(* IEC 61131-3 sources: plc-st-coding-agent/progress/evidence/f14_v13_self_20261113/jobs/custom_deepseek-v4pro (part 4) *)

(* ---- public-medium-02.raw_candidate_01.st ---- *)
TYPE ST_AnalogChannel :
STRUCT
    enable : BOOL;
    hiLIM : REAL;
    loLIM : REAL;
    bipolar : BOOL;
    measuringMode : INT;
    retVal : WORD;
    outputValue : REAL;
END_STRUCT
END_TYPE

(* ENGINEERING_CONTRACT
   Loop count: count limited to 0..min(array lengths); ordinal start at each array lower bound (PUB001).
   channels[].retVal: activated on enabled scan; invalid mode -> 16#8001, invalid limits -> 16#8002,
   success -> 0 (PUB006, PUB007, PUB008).
   channels[].outputValue: written only on successful conversion; mode 0 linear scaling,
   mode 1 /10, mode 2 /100 (PUB003, PUB004, PUB005).
   Disabled channels retain prior retVal/outputValue (unspecified retention interpretation).
*)

(* CONTRACT_RULES [] *)

FUNCTION_BLOCK AnalogBatchProcessing
VAR_INPUT
    count : DINT;
END_VAR
VAR_IN_OUT
    analogValues : ARRAY[*] OF INT;
    channels : ARRAY[*] OF ST_AnalogChannel;
END_VAR
VAR
    local_i : DINT;
    local_n : DINT;
    local_analog_idx : DINT;
    local_channel_idx : DINT;
    local_raw : INT;
    local_mode : INT;
    local_min_len : DINT;
    local_ch_len : DINT;
    local_raw_min : REAL;
    local_raw_max : REAL;
    local_span_raw : REAL;
    local_ratio : REAL;
END_VAR

local_n := count;
IF local_n < 0 THEN
    local_n := 0;
END_IF;

local_min_len := UPPER_BOUND(analogValues, 1) - LOWER_BOUND(analogValues, 1) + 1;
local_ch_len := UPPER_BOUND(channels, 1) - LOWER_BOUND(channels, 1) + 1;
IF local_min_len > local_ch_len THEN
    local_min_len := local_ch_len;
END_IF;
IF local_n > local_min_len THEN
    local_n := local_min_len;
END_IF;

IF local_n > 0 THEN
    FOR local_i := 0 TO local_n - 1 DO
        local_analog_idx := LOWER_BOUND(analogValues, 1) + local_i;
        local_channel_idx := LOWER_BOUND(channels, 1) + local_i;

        IF channels[local_channel_idx].enable THEN
            local_mode := channels[local_channel_idx].measuringMode;

            IF (local_mode <> 0) AND (local_mode <> 1) AND (local_mode <> 2) THEN
                channels[local_channel_idx].retVal := 16#8001;
                (* skip conversion: outputValue unchanged *)
            ELSIF channels[local_channel_idx].hiLIM <= channels[local_channel_idx].loLIM THEN
                channels[local_channel_idx].retVal := 16#8002;
                (* skip conversion: outputValue unchanged *)
            ELSE
                channels[local_channel_idx].retVal := 0;
                CASE local_mode OF
                    0:
                        local_raw := analogValues[local_analog_idx];
                        IF channels[local_channel_idx].bipolar THEN
                            local_raw_min := -27648.0;
                            local_raw_max := 27648.0;
                        ELSE
                            local_raw_min := 0.0;
                            local_raw_max := 27648.0;
                        END_IF;

                        local_span_raw := local_raw_max - local_raw_min;
                        local_ratio := (TO_REAL(local_raw) - local_raw_min) / local_span_raw;
                        channels[local_channel_idx].outputValue := channels[local_channel_idx].loLIM
                            + local_ratio * (channels[local_channel_idx].hiLIM - channels[local_channel_idx].loLIM);

                    1:
                        channels[local_channel_idx].outputValue := TO_REAL(analogValues[local_analog_idx]) / 10.0;

                    2:
                        channels[local_channel_idx].outputValue := TO_REAL(analogValues[local_analog_idx]) / 100.0;
                END_CASE;
            END_IF;
        ELSE
            (* disabled: no writes to retVal or outputValue *)
        END_IF;
    END_FOR;
END_IF;

(* ---- public-medium-02.raw_candidate_02.st ---- *)
TYPE ST_AnalogChannel :
STRUCT
    enable : BOOL;
    hiLIM : REAL;
    loLIM : REAL;
    bipolar : BOOL;
    measuringMode : INT;
    retVal : WORD;
    outputValue : REAL;
END_STRUCT
END_TYPE;

(* ENGINEERING_CONTRACT
   Loop count: count limited to 0..min(array lengths); ordinal start at each array lower bound (PUB001).
   channels[].retVal: activated on enabled scan; invalid mode -> 16#8001, invalid limits -> 16#8002,
   success -> 0 (PUB006, PUB007, PUB008).
   channels[].outputValue: written only on successful conversion; mode 0 linear scaling,
   mode 1 /10, mode 2 /100 (PUB003, PUB004, PUB005).
   Disabled channels retain prior retVal/outputValue (unspecified retention interpretation).
*)

(* CONTRACT_RULES [] *)

FUNCTION_BLOCK AnalogBatchProcessing
VAR_INPUT
    count : DINT;
END_VAR
VAR_IN_OUT
    analogValues : ARRAY[*] OF INT;
    channels : ARRAY[*] OF ST_AnalogChannel;
END_VAR
VAR
    local_i : DINT;
    local_n : DINT;
    local_analog_idx : DINT;
    local_channel_idx : DINT;
    local_raw : INT;
    local_mode : INT;
    local_min_len : DINT;
    local_ch_len : DINT;
    local_raw_min : REAL;
    local_raw_max : REAL;
    local_span_raw : REAL;
    local_ratio : REAL;
END_VAR

local_n := count;
IF local_n < 0 THEN
    local_n := 0;
END_IF;

local_min_len := UPPER_BOUND(analogValues, 1) - LOWER_BOUND(analogValues, 1) + 1;
local_ch_len := UPPER_BOUND(channels, 1) - LOWER_BOUND(channels, 1) + 1;
IF local_min_len > local_ch_len THEN
    local_min_len := local_ch_len;
END_IF;
IF local_n > local_min_len THEN
    local_n := local_min_len;
END_IF;

IF local_n > 0 THEN
    FOR local_i := 0 TO local_n - 1 DO
        local_analog_idx := LOWER_BOUND(analogValues, 1) + local_i;
        local_channel_idx := LOWER_BOUND(channels, 1) + local_i;

        IF channels[local_channel_idx].enable THEN
            local_mode := channels[local_channel_idx].measuringMode;

            IF (local_mode <> 0) AND (local_mode <> 1) AND (local_mode <> 2) THEN
                channels[local_channel_idx].retVal := 16#8001;
                (* skip conversion: outputValue unchanged *)
            ELSIF channels[local_channel_idx].hiLIM <= channels[local_channel_idx].loLIM THEN
                channels[local_channel_idx].retVal := 16#8002;
                (* skip conversion: outputValue unchanged *)
            ELSE
                channels[local_channel_idx].retVal := 0;
                CASE local_mode OF
                    0:
                        local_raw := analogValues[local_analog_idx];
                        IF channels[local_channel_idx].bipolar THEN
                            local_raw_min := -27648.0;
                            local_raw_max := 27648.0;
                        ELSE
                            local_raw_min := 0.0;
                            local_raw_max := 27648.0;
                        END_IF;

                        local_span_raw := local_raw_max - local_raw_min;
                        local_ratio := (TO_REAL(local_raw) - local_raw_min) / local_span_raw;
                        channels[local_channel_idx].outputValue := channels[local_channel_idx].loLIM
                            + local_ratio * (channels[local_channel_idx].hiLIM - channels[local_channel_idx].loLIM);

                    1:
                        channels[local_channel_idx].outputValue := TO_REAL(analogValues[local_analog_idx]) / 10.0;

                    2:
                        channels[local_channel_idx].outputValue := TO_REAL(analogValues[local_analog_idx]) / 100.0;
                END_CASE;
            END_IF;
        ELSE
            (* disabled: no writes to retVal or outputValue *)
        END_IF;
    END_FOR;
END_IF;

END_FUNCTION_BLOCK

(* ---- public-medium-02.raw_candidate_03.st ---- *)
TYPE ST_AnalogChannel :
STRUCT
    enable : BOOL;
    hiLIM : REAL;
    loLIM : REAL;
    bipolar : BOOL;
    measuringMode : INT;
    retVal : WORD;
    outputValue : REAL;
END_STRUCT
END_TYPE

(* ENGINEERING_CONTRACT
   Loop count: count limited to 0..min(array lengths); ordinal start at each array lower bound (PUB001).
   channels[].retVal: activated on enabled scan; invalid mode -> 16#8001, invalid limits -> 16#8002,
   success -> 0 (PUB006, PUB007, PUB008).
   channels[].outputValue: written only on successful conversion; mode 0 linear scaling,
   mode 1 /10, mode 2 /100 (PUB003, PUB004, PUB005).
   Disabled channels retain prior retVal/outputValue (unspecified retention interpretation).
*)

(* CONTRACT_RULES [] *)

FUNCTION_BLOCK AnalogBatchProcessing
VAR_INPUT
    count : DINT;
END_VAR
VAR_IN_OUT
    analogValues : ARRAY[*] OF INT;
    channels : ARRAY[*] OF ST_AnalogChannel;
END_VAR
VAR
    local_i : DINT;
    local_n : DINT;
    local_analog_idx : DINT;
    local_channel_idx : DINT;
    local_raw : INT;
    local_mode : INT;
    local_min_len : DINT;
    local_ch_len : DINT;
    local_raw_min : REAL;
    local_raw_max : REAL;
    local_span_raw : REAL;
    local_ratio : REAL;
END_VAR

local_n := count;
IF local_n < 0 THEN
    local_n := 0;
END_IF;

local_min_len := UPPER_BOUND(analogValues, 1) - LOWER_BOUND(analogValues, 1) + 1;
local_ch_len := UPPER_BOUND(channels, 1) - LOWER_BOUND(channels, 1) + 1;
IF local_min_len > local_ch_len THEN
    local_min_len := local_ch_len;
END_IF;
IF local_n > local_min_len THEN
    local_n := local_min_len;
END_IF;

IF local_n > 0 THEN
    FOR local_i := 0 TO local_n - 1 DO
        local_analog_idx := LOWER_BOUND(analogValues, 1) + local_i;
        local_channel_idx := LOWER_BOUND(channels, 1) + local_i;

        IF channels[local_channel_idx].enable THEN
            local_mode := channels[local_channel_idx].measuringMode;

            IF (local_mode <> 0) AND (local_mode <> 1) AND (local_mode <> 2) THEN
                channels[local_channel_idx].retVal := 16#8001;
                (* skip conversion: outputValue unchanged *)
            ELSIF channels[local_channel_idx].hiLIM <= channels[local_channel_idx].loLIM THEN
                channels[local_channel_idx].retVal := 16#8002;
                (* skip conversion: outputValue unchanged *)
            ELSE
                channels[local_channel_idx].retVal := 0;
                CASE local_mode OF
                    0:
                        local_raw := analogValues[local_analog_idx];
                        IF channels[local_channel_idx].bipolar THEN
                            local_raw_min := -27648.0;
                            local_raw_max := 27648.0;
                        ELSE
                            local_raw_min := 0.0;
                            local_raw_max := 27648.0;
                        END_IF;

                        local_span_raw := local_raw_max - local_raw_min;
                        local_ratio := (TO_REAL(local_raw) - local_raw_min) / local_span_raw;
                        channels[local_channel_idx].outputValue := channels[local_channel_idx].loLIM
                            + local_ratio * (channels[local_channel_idx].hiLIM - channels[local_channel_idx].loLIM);

                    1:
                        channels[local_channel_idx].outputValue := TO_REAL(analogValues[local_analog_idx]) / 10.0;

                    2:
                        channels[local_channel_idx].outputValue := TO_REAL(analogValues[local_analog_idx]) / 100.0;
                END_CASE;
            END_IF;
        ELSE
            (* disabled: no writes to retVal or outputValue *)
        END_IF;
    END_FOR;
END_IF;

END_FUNCTION_BLOCK

(* ---- public-medium-03.candidate_01.st ---- *)
(* ENGINEERING_CONTRACT
- average: stored LREAL; updated on valid acquisition; reset or invalid window clears it to 0.0.
- windowSizeReached: FALSE until count >= windowSize; retained until reset or invalid window.
- error/status: combinational invalid windowSize (1..100 inclusive); otherwise clear/zero.
- Priority: invalid window first, reset second, acquisition last (reset priority chosen).
- cyclicExecution TRUE ignores trigger edges for extra samples (PUB001/2).
- trigger edge is evaluated only from previous scan raw trigger state.
- Same-scan: validate window, detect window-size change, reset, acquire, update average.
*)
(* CONTRACT_RULES [] *)
FUNCTION_BLOCK FB
VAR_INPUT
    cyclicExecution : BOOL;
    trigger : BOOL;
    value : LREAL;
    windowSize : INT;
    reset : BOOL;
END_VAR
VAR_OUTPUT
    average : LREAL;
    windowSizeReached : BOOL;
    error : BOOL;
    status : WORD;
END_VAR
VAR
    tmp_buffer : ARRAY[0..99] OF LREAL;
    tmp_count : INT := 0;
    tmp_index : INT := 0;
    tmp_sum : LREAL := 0.0;
    tmp_previousTrigger : BOOL := FALSE;
    tmp_windowSize : INT := 0;
END_VAR

IF (windowSize < 1) OR (windowSize > 100) THEN
    error := TRUE;
    status := WORD#16#8200;
    windowSizeReached := FALSE;
    average := 0.0;
    tmp_count := 0;
    tmp_index := 0;
    tmp_sum := 0.0;
    tmp_windowSize := windowSize;
ELSE
    error := FALSE;
    status := WORD#16#0000;

    IF tmp_windowSize <> windowSize THEN
        tmp_count := 0;
        tmp_index := 0;
        tmp_sum := 0.0;
        windowSizeReached := FALSE;
        average := 0.0;
        tmp_windowSize := windowSize;
    END_IF;

    IF reset THEN
        tmp_count := 0;
        tmp_index := 0;
        tmp_sum := 0.0;
        windowSizeReached := FALSE;
        average := 0.0;
    ELSE
        IF cyclicExecution OR (trigger AND NOT tmp_previousTrigger) THEN
            IF tmp_count < windowSize THEN
                tmp_count := tmp_count + 1;
                tmp_sum := tmp_sum + value;
                tmp_buffer[tmp_index] := value;
                tmp_index := tmp_index + 1;
                IF tmp_index >= windowSize THEN
                    tmp_index := 0;
                END_IF;
            ELSE
                tmp_sum := tmp_sum - tmp_buffer[tmp_index] + value;
                tmp_buffer[tmp_index] := value;
                tmp_index := tmp_index + 1;
                IF tmp_index >= windowSize THEN
                    tmp_index := 0;
                END_IF;
            END_IF;

            average := tmp_sum / INT_TO_LREAL(tmp_count);
            windowSizeReached := tmp_count >= windowSize;
        END_IF;
    END_IF;
END_IF;

tmp_previousTrigger := trigger;

(* ---- public-medium-03.candidate_02.st ---- *)
(* ENGINEERING_CONTRACT
- average: stored LREAL; updated on valid acquisition; reset or invalid window clears it to 0.0.
- windowSizeReached: FALSE until count >= windowSize; retained until reset or invalid window.
- error/status: combinational invalid windowSize (1..100 inclusive); otherwise clear/zero.
- Priority: invalid window first, reset second, acquisition last (reset priority chosen).
- cyclicExecution TRUE ignores trigger edges for extra samples (PUB001/2).
- trigger edge is evaluated only from previous scan raw trigger state.
- Same-scan: validate window, detect window-size change, reset, acquire, update average.
*)
(* CONTRACT_RULES [] *)
FUNCTION_BLOCK FB
VAR_INPUT
    cyclicExecution : BOOL;
    trigger : BOOL;
    value : LREAL;
    windowSize : INT;
    reset : BOOL;
END_VAR
VAR_OUTPUT
    average : LREAL;
    windowSizeReached : BOOL;
    error : BOOL;
    status : WORD;
END_VAR
VAR
    tmp_buffer : ARRAY[0..99] OF LREAL;
    tmp_count : INT := 0;
    tmp_index : INT := 0;
    tmp_sum : LREAL := 0.0;
    tmp_previousTrigger : BOOL := FALSE;
    tmp_windowSize : INT := 0;
END_VAR

IF (windowSize < 1) OR (windowSize > 100) THEN
    error := TRUE;
    status := WORD#16#8200;
    windowSizeReached := FALSE;
    average := 0.0;
    tmp_count := 0;
    tmp_index := 0;
    tmp_sum := 0.0;
    tmp_windowSize := windowSize;
ELSE
    error := FALSE;
    status := WORD#16#0000;

    IF tmp_windowSize <> windowSize THEN
        tmp_count := 0;
        tmp_index := 0;
        tmp_sum := 0.0;
        windowSizeReached := FALSE;
        average := 0.0;
        tmp_windowSize := windowSize;
    END_IF;

    IF reset THEN
        tmp_count := 0;
        tmp_index := 0;
        tmp_sum := 0.0;
        windowSizeReached := FALSE;
        average := 0.0;
    ELSE
        IF cyclicExecution OR (trigger AND NOT tmp_previousTrigger) THEN
            IF tmp_count < windowSize THEN
                tmp_count := tmp_count + 1;
                tmp_sum := tmp_sum + value;
                tmp_buffer[tmp_index] := value;
                tmp_index := tmp_index + 1;
                IF tmp_index >= windowSize THEN
                    tmp_index := 0;
                END_IF;
            ELSE
                tmp_sum := tmp_sum - tmp_buffer[tmp_index] + value;
                tmp_buffer[tmp_index] := value;
                tmp_index := tmp_index + 1;
                IF tmp_index >= windowSize THEN
                    tmp_index := 0;
                END_IF;
            END_IF;

            average := tmp_sum / INT_TO_LREAL(tmp_count);
            windowSizeReached := tmp_count >= windowSize;
        END_IF;
    END_IF;
END_IF;

tmp_previousTrigger := trigger;
END_FUNCTION_BLOCK

(* ---- public-medium-03.patch_base_02.st ---- *)
(* ENGINEERING_CONTRACT
- average: stored LREAL; updated on valid acquisition; reset or invalid window clears it to 0.0.
- windowSizeReached: FALSE until count >= windowSize; retained until reset or invalid window.
- error/status: combinational invalid windowSize (1..100 inclusive); otherwise clear/zero.
- Priority: invalid window first, reset second, acquisition last (reset priority chosen).
- cyclicExecution TRUE ignores trigger edges for extra samples (PUB001/2).
- trigger edge is evaluated only from previous scan raw trigger state.
- Same-scan: validate window, detect window-size change, reset, acquire, update average.
*)
(* CONTRACT_RULES [] *)
FUNCTION_BLOCK FB
VAR_INPUT
    cyclicExecution : BOOL;
    trigger : BOOL;
    value : LREAL;
    windowSize : INT;
    reset : BOOL;
END_VAR
VAR_OUTPUT
    average : LREAL;
    windowSizeReached : BOOL;
    error : BOOL;
    status : WORD;
END_VAR
VAR
    tmp_buffer : ARRAY[0..99] OF LREAL;
    tmp_count : INT := 0;
    tmp_index : INT := 0;
    tmp_sum : LREAL := 0.0;
    tmp_previousTrigger : BOOL := FALSE;
    tmp_windowSize : INT := 0;
END_VAR

IF (windowSize < 1) OR (windowSize > 100) THEN
    error := TRUE;
    status := WORD#16#8200;
    windowSizeReached := FALSE;
    average := 0.0;
    tmp_count := 0;
    tmp_index := 0;
    tmp_sum := 0.0;
    tmp_windowSize := windowSize;
ELSE
    error := FALSE;
    status := WORD#16#0000;

    IF tmp_windowSize <> windowSize THEN
        tmp_count := 0;
        tmp_index := 0;
        tmp_sum := 0.0;
        windowSizeReached := FALSE;
        average := 0.0;
        tmp_windowSize := windowSize;
    END_IF;

    IF reset THEN
        tmp_count := 0;
        tmp_index := 0;
        tmp_sum := 0.0;
        windowSizeReached := FALSE;
        average := 0.0;
    ELSE
        IF cyclicExecution OR (trigger AND NOT tmp_previousTrigger) THEN
            IF tmp_count < windowSize THEN
                tmp_count := tmp_count + 1;
                tmp_sum := tmp_sum + value;
                tmp_buffer[tmp_index] := value;
                tmp_index := tmp_index + 1;
                IF tmp_index >= windowSize THEN
                    tmp_index := 0;
                END_IF;
            ELSE
                tmp_sum := tmp_sum - tmp_buffer[tmp_index] + value;
                tmp_buffer[tmp_index] := value;
                tmp_index := tmp_index + 1;
                IF tmp_index >= windowSize THEN
                    tmp_index := 0;
                END_IF;
            END_IF;

            average := tmp_sum / INT_TO_LREAL(tmp_count);
            windowSizeReached := tmp_count >= windowSize;
        END_IF;
    END_IF;
END_IF;

tmp_previousTrigger := trigger;

(* ---- public-medium-03.raw_candidate_01.st ---- *)
(* ENGINEERING_CONTRACT
- average: stored LREAL; updated on valid acquisition; reset or invalid window clears it to 0.0.
- windowSizeReached: FALSE until count >= windowSize; retained until reset or invalid window.
- error/status: combinational invalid windowSize (1..100 inclusive); otherwise clear/zero.
- Priority: invalid window first, reset second, acquisition last (reset priority chosen).
- cyclicExecution TRUE ignores trigger edges for extra samples (PUB001/2).
- trigger edge is evaluated only from previous scan raw trigger state.
- Same-scan: validate window, detect window-size change, reset, acquire, update average.
*)
(* CONTRACT_RULES [] *)
FUNCTION_BLOCK FB
VAR_INPUT
    cyclicExecution : BOOL;
    trigger : BOOL;
    value : LREAL;
    windowSize : INT;
    reset : BOOL;
END_VAR
VAR_OUTPUT
    average : LREAL;
    windowSizeReached : BOOL;
    error : BOOL;
    status : WORD;
END_VAR
VAR
    tmp_buffer : ARRAY[0..99] OF LREAL;
    tmp_count : INT := 0;
    tmp_index : INT := 0;
    tmp_sum : LREAL := 0.0;
    tmp_previousTrigger : BOOL := FALSE;
    tmp_windowSize : INT := 0;
END_VAR

IF (windowSize < 1) OR (windowSize > 100) THEN
    error := TRUE;
    status := WORD#16#8200;
    windowSizeReached := FALSE;
    average := 0.0;
    tmp_count := 0;
    tmp_index := 0;
    tmp_sum := 0.0;
    tmp_windowSize := windowSize;
ELSE
    error := FALSE;
    status := WORD#16#0000;

    IF tmp_windowSize <> windowSize THEN
        tmp_count := 0;
        tmp_index := 0;
        tmp_sum := 0.0;
        windowSizeReached := FALSE;
        average := 0.0;
        tmp_windowSize := windowSize;
    END_IF;

    IF reset THEN
        tmp_count := 0;
        tmp_index := 0;
        tmp_sum := 0.0;
        windowSizeReached := FALSE;
        average := 0.0;
    ELSE
        IF cyclicExecution OR (trigger AND NOT tmp_previousTrigger) THEN
            IF tmp_count < windowSize THEN
                tmp_count := tmp_count + 1;
                tmp_sum := tmp_sum + value;
                tmp_buffer[tmp_index] := value;
                tmp_index := tmp_index + 1;
                IF tmp_index >= windowSize THEN
                    tmp_index := 0;
                END_IF;
            ELSE
                tmp_sum := tmp_sum - tmp_buffer[tmp_index] + value;
                tmp_buffer[tmp_index] := value;
                tmp_index := tmp_index + 1;
                IF tmp_index >= windowSize THEN
                    tmp_index := 0;
                END_IF;
            END_IF;

            average := tmp_sum / INT_TO_LREAL(tmp_count);
            windowSizeReached := tmp_count >= windowSize;
        END_IF;
    END_IF;
END_IF;

tmp_previousTrigger := trigger;

(* ---- public-medium-03.raw_candidate_02.st ---- *)
(* ENGINEERING_CONTRACT
- average: stored LREAL; updated on valid acquisition; reset or invalid window clears it to 0.0.
- windowSizeReached: FALSE until count >= windowSize; retained until reset or invalid window.
- error/status: combinational invalid windowSize (1..100 inclusive); otherwise clear/zero.
- Priority: invalid window first, reset second, acquisition last (reset priority chosen).
- cyclicExecution TRUE ignores trigger edges for extra samples (PUB001/2).
- trigger edge is evaluated only from previous scan raw trigger state.
- Same-scan: validate window, detect window-size change, reset, acquire, update average.
*)
(* CONTRACT_RULES [] *)
FUNCTION_BLOCK FB
VAR_INPUT
    cyclicExecution : BOOL;
    trigger : BOOL;
    value : LREAL;
    windowSize : INT;
    reset : BOOL;
END_VAR
VAR_OUTPUT
    average : LREAL;
    windowSizeReached : BOOL;
    error : BOOL;
    status : WORD;
END_VAR
VAR
    tmp_buffer : ARRAY[0..99] OF LREAL;
    tmp_count : INT := 0;
    tmp_index : INT := 0;
    tmp_sum : LREAL := 0.0;
    tmp_previousTrigger : BOOL := FALSE;
    tmp_windowSize : INT := 0;
END_VAR

IF (windowSize < 1) OR (windowSize > 100) THEN
    error := TRUE;
    status := WORD#16#8200;
    windowSizeReached := FALSE;
    average := 0.0;
    tmp_count := 0;
    tmp_index := 0;
    tmp_sum := 0.0;
    tmp_windowSize := windowSize;
ELSE
    error := FALSE;
    status := WORD#16#0000;

    IF tmp_windowSize <> windowSize THEN
        tmp_count := 0;
        tmp_index := 0;
        tmp_sum := 0.0;
        windowSizeReached := FALSE;
        average := 0.0;
        tmp_windowSize := windowSize;
    END_IF;

    IF reset THEN
        tmp_count := 0;
        tmp_index := 0;
        tmp_sum := 0.0;
        windowSizeReached := FALSE;
        average := 0.0;
    ELSE
        IF cyclicExecution OR (trigger AND NOT tmp_previousTrigger) THEN
            IF tmp_count < windowSize THEN
                tmp_count := tmp_count + 1;
                tmp_sum := tmp_sum + value;
                tmp_buffer[tmp_index] := value;
                tmp_index := tmp_index + 1;
                IF tmp_index >= windowSize THEN
                    tmp_index := 0;
                END_IF;
            ELSE
                tmp_sum := tmp_sum - tmp_buffer[tmp_index] + value;
                tmp_buffer[tmp_index] := value;
                tmp_index := tmp_index + 1;
                IF tmp_index >= windowSize THEN
                    tmp_index := 0;
                END_IF;
            END_IF;

            average := tmp_sum / INT_TO_LREAL(tmp_count);
            windowSizeReached := tmp_count >= windowSize;
        END_IF;
    END_IF;
END_IF;

tmp_previousTrigger := trigger;
END_FUNCTION_BLOCK

(* ---- public-medium-04.candidate_01.st ---- *)
FUNCTION_BLOCK FB_TemperatureControl
VAR_INPUT
    TemperatureSensorInput : REAL;
    SetTemperature : REAL;
END_VAR
VAR_OUTPUT
    CurrentTemperature : REAL;
    SetTempDisplay : REAL;
    HeaterStatus : BOOL;
    OverheatProtection : BOOL;
    HeaterOutput : BOOL;
END_VAR
VAR
    local_OverheatActive : BOOL := FALSE;
    local_SensorFault : BOOL;
    local_DesiredHeater : BOOL;
    tmp_HeaterOnTimer : TON;
    tmp_CooldownTimer : TON;
END_VAR

(* ENGINEERING_CONTRACT
   CurrentTemperature/SetTempDisplay: mirror inputs every scan; no retention.
   HeaterOutput: ON only when sensor OK, protection inactive and temp < set (PUB003).
     OFF when temp >= set (PUB004; equality unspecified, implemented OFF).
   Sensor fault (input < 0 or > 100) forces OFF (PUB007).
   OverheatProtection: set when HeaterOutput continuously TRUE > 5000 ms via TON (PUB005).
     Retained TRUE until 3 s cooldown TON completes; then clears automatically (PUB005).
   Same-scan priority: sensor fault and overheat protection override normal compare (PUB005/PUB007).
   HeaterStatus mirrors final HeaterOutput; temperatures in deg C; thresholds strict.
*)
(* CONTRACT_RULES [] *)

CurrentTemperature := TemperatureSensorInput;
SetTempDisplay := SetTemperature;

local_SensorFault := (TemperatureSensorInput < 0.0) OR (TemperatureSensorInput > 100.0);

tmp_CooldownTimer(IN := local_OverheatActive, PT := T#3S);
IF tmp_CooldownTimer.Q THEN
    local_OverheatActive := FALSE;
END_IF;

IF local_SensorFault THEN
    local_DesiredHeater := FALSE;
ELSIF local_OverheatActive THEN
    local_DesiredHeater := FALSE;
ELSE
    IF TemperatureSensorInput < SetTemperature THEN
        local_DesiredHeater := TRUE;
    ELSE
        local_DesiredHeater := FALSE;
    END_IF;
END_IF;

HeaterOutput := local_DesiredHeater;

tmp_HeaterOnTimer(IN := HeaterOutput, PT := T#5001MS);
IF tmp_HeaterOnTimer.Q THEN
    local_OverheatActive := TRUE;
    HeaterOutput := FALSE;
END_IF;

HeaterStatus := HeaterOutput;
OverheatProtection := local_OverheatActive;
END_FUNCTION_BLOCK

(* ---- public-medium-04.candidate_02.st ---- *)
FUNCTION_BLOCK FB_TemperatureControl
VAR_INPUT
    TemperatureSensorInput : REAL;
    SetTemperature : REAL;
END_VAR
VAR_OUTPUT
    CurrentTemperature : REAL;
    SetTempDisplay : REAL;
    HeaterStatus : BOOL;
    OverheatProtection : BOOL;
    HeaterOutput : BOOL;
END_VAR
VAR
    local_OverheatActive : BOOL := FALSE;
    local_SensorFault : BOOL;
    local_DesiredHeater : BOOL;
    tmp_HeaterOnTimer : TON;
    tmp_CooldownTimer : TON;
END_VAR

(* ENGINEERING_CONTRACT
   CurrentTemperature/SetTempDisplay: mirror inputs every scan; no retention.
   HeaterOutput: ON only when sensor OK, protection inactive and temp < set (PUB003).
     OFF when temp >= set (PUB004; equality unspecified, implemented OFF).
   Sensor fault (input < 0 or > 100) forces OFF (PUB007).
   OverheatProtection: set when HeaterOutput continuously TRUE > 5000 ms via TON (PUB005).
     Retained TRUE until 3 s cooldown TON completes; then clears automatically (PUB005).
   Same-scan priority: sensor fault and overheat protection override normal compare (PUB005/PUB007).
   HeaterStatus mirrors final HeaterOutput; temperatures in deg C; thresholds strict.
*)
(* CONTRACT_RULES [] *)

CurrentTemperature := TemperatureSensorInput;
SetTempDisplay := SetTemperature;

local_SensorFault := (TemperatureSensorInput < 0.0) OR (TemperatureSensorInput > 100.0);

IF local_SensorFault OR local_OverheatActive THEN
    local_DesiredHeater := FALSE;
ELSIF TemperatureSensorInput < SetTemperature THEN
    local_DesiredHeater := TRUE;
ELSE
    local_DesiredHeater := FALSE;
END_IF;

HeaterOutput := local_DesiredHeater;

tmp_HeaterOnTimer(IN := HeaterOutput, PT := T#5001MS);
IF tmp_HeaterOnTimer.Q THEN
    local_OverheatActive := TRUE;
    HeaterOutput := FALSE;
END_IF;

tmp_CooldownTimer(IN := local_OverheatActive, PT := T#3S);
IF tmp_CooldownTimer.Q THEN
    local_OverheatActive := FALSE;
    IF local_SensorFault THEN
        HeaterOutput := FALSE;
    ELSIF TemperatureSensorInput < SetTemperature THEN
        HeaterOutput := TRUE;
    ELSE
        HeaterOutput := FALSE;
    END_IF;
    tmp_HeaterOnTimer(IN := HeaterOutput, PT := T#5001MS);
END_IF;

HeaterStatus := HeaterOutput;
OverheatProtection := local_OverheatActive;
END_FUNCTION_BLOCK

(* ---- public-medium-04.patch_base_02.st ---- *)
FUNCTION_BLOCK FB_TemperatureControl
VAR_INPUT
    TemperatureSensorInput : REAL;
    SetTemperature : REAL;
END_VAR
VAR_OUTPUT
    CurrentTemperature : REAL;
    SetTempDisplay : REAL;
    HeaterStatus : BOOL;
    OverheatProtection : BOOL;
    HeaterOutput : BOOL;
END_VAR
VAR
    local_OverheatActive : BOOL := FALSE;
    local_SensorFault : BOOL;
    local_DesiredHeater : BOOL;
    tmp_HeaterOnTimer : TON;
    tmp_CooldownTimer : TON;
END_VAR

(* ENGINEERING_CONTRACT
   CurrentTemperature/SetTempDisplay: mirror inputs every scan; no retention.
   HeaterOutput: ON only when sensor OK, protection inactive and temp < set (PUB003).
     OFF when temp >= set (PUB004; equality unspecified, implemented OFF).
   Sensor fault (input < 0 or > 100) forces OFF (PUB007).
   OverheatProtection: set when HeaterOutput continuously TRUE > 5000 ms via TON (PUB005).
     Retained TRUE until 3 s cooldown TON completes; then clears automatically (PUB005).
   Same-scan priority: sensor fault and overheat protection override normal compare (PUB005/PUB007).
   HeaterStatus mirrors final HeaterOutput; temperatures in deg C; thresholds strict.
*)
(* CONTRACT_RULES [] *)

CurrentTemperature := TemperatureSensorInput;
SetTempDisplay := SetTemperature;

local_SensorFault := (TemperatureSensorInput < 0.0) OR (TemperatureSensorInput > 100.0);

tmp_CooldownTimer(IN := local_OverheatActive, PT := T#3S);
IF tmp_CooldownTimer.Q THEN
    local_OverheatActive := FALSE;
END_IF;

IF local_SensorFault THEN
    local_DesiredHeater := FALSE;
ELSIF local_OverheatActive THEN
    local_DesiredHeater := FALSE;
ELSE
    IF TemperatureSensorInput < SetTemperature THEN
        local_DesiredHeater := TRUE;
    ELSE
        local_DesiredHeater := FALSE;
    END_IF;
END_IF;

HeaterOutput := local_DesiredHeater;

tmp_HeaterOnTimer(IN := HeaterOutput, PT := T#5001MS);
IF tmp_HeaterOnTimer.Q THEN
    local_OverheatActive := TRUE;
    HeaterOutput := FALSE;
END_IF;

HeaterStatus := HeaterOutput;
OverheatProtection := local_OverheatActive;
END_FUNCTION_BLOCK

(* ---- public-medium-04.raw_candidate_01.st ---- *)
FUNCTION_BLOCK FB_TemperatureControl
VAR_INPUT
    TemperatureSensorInput : REAL;
    SetTemperature : REAL;
END_VAR
VAR_OUTPUT
    CurrentTemperature : REAL;
    SetTempDisplay : REAL;
    HeaterStatus : BOOL;
    OverheatProtection : BOOL;
    HeaterOutput : BOOL;
END_VAR
VAR
    local_OverheatActive : BOOL := FALSE;
    local_SensorFault : BOOL;
    local_DesiredHeater : BOOL;
    tmp_HeaterOnTimer : TON;
    tmp_CooldownTimer : TON;
END_VAR

(* ENGINEERING_CONTRACT
   CurrentTemperature/SetTempDisplay: mirror inputs every scan; no retention.
   HeaterOutput: ON only when sensor OK, protection inactive and temp < set (PUB003).
     OFF when temp >= set (PUB004; equality unspecified, implemented OFF).
   Sensor fault (input < 0 or > 100) forces OFF (PUB007).
   OverheatProtection: set when HeaterOutput continuously TRUE > 5000 ms via TON (PUB005).
     Retained TRUE until 3 s cooldown TON completes; then clears automatically (PUB005).
   Same-scan priority: sensor fault and overheat protection override normal compare (PUB005/PUB007).
   HeaterStatus mirrors final HeaterOutput; temperatures in deg C; thresholds strict.
*)
(* CONTRACT_RULES [] *)

CurrentTemperature := TemperatureSensorInput;
SetTempDisplay := SetTemperature;

local_SensorFault := (TemperatureSensorInput < 0.0) OR (TemperatureSensorInput > 100.0);

tmp_CooldownTimer(IN := local_OverheatActive, PT := T#3S);
IF tmp_CooldownTimer.Q THEN
    local_OverheatActive := FALSE;
END_IF;

IF local_SensorFault THEN
    local_DesiredHeater := FALSE;
ELSIF local_OverheatActive THEN
    local_DesiredHeater := FALSE;
ELSE
    IF TemperatureSensorInput < SetTemperature THEN
        local_DesiredHeater := TRUE;
    ELSE
        local_DesiredHeater := FALSE;
    END_IF;
END_IF;

HeaterOutput := local_DesiredHeater;

tmp_HeaterOnTimer(IN := HeaterOutput, PT := T#5001MS);
IF tmp_HeaterOnTimer.Q THEN
    local_OverheatActive := TRUE;
    HeaterOutput := FALSE;
END_IF;

HeaterStatus := HeaterOutput;
OverheatProtection := local_OverheatActive;
END_FUNCTION_BLOCK

(* ---- public-medium-04.raw_candidate_02.st ---- *)
FUNCTION_BLOCK FB_TemperatureControl
VAR_INPUT
    TemperatureSensorInput : REAL;
    SetTemperature : REAL;
END_VAR
VAR_OUTPUT
    CurrentTemperature : REAL;
    SetTempDisplay : REAL;
    HeaterStatus : BOOL;
    OverheatProtection : BOOL;
    HeaterOutput : BOOL;
END_VAR
VAR
    local_OverheatActive : BOOL := FALSE;
    local_SensorFault : BOOL;
    local_DesiredHeater : BOOL;
    tmp_HeaterOnTimer : TON;
    tmp_CooldownTimer : TON;
END_VAR

(* ENGINEERING_CONTRACT
   CurrentTemperature/SetTempDisplay: mirror inputs every scan; no retention.
   HeaterOutput: ON only when sensor OK, protection inactive and temp < set (PUB003).
     OFF when temp >= set (PUB004; equality unspecified, implemented OFF).
   Sensor fault (input < 0 or > 100) forces OFF (PUB007).
   OverheatProtection: set when HeaterOutput continuously TRUE > 5000 ms via TON (PUB005).
     Retained TRUE until 3 s cooldown TON completes; then clears automatically (PUB005).
   Same-scan priority: sensor fault and overheat protection override normal compare (PUB005/PUB007).
   HeaterStatus mirrors final HeaterOutput; temperatures in deg C; thresholds strict.
*)
(* CONTRACT_RULES [] *)

CurrentTemperature := TemperatureSensorInput;
SetTempDisplay := SetTemperature;

local_SensorFault := (TemperatureSensorInput < 0.0) OR (TemperatureSensorInput > 100.0);

IF local_SensorFault OR local_OverheatActive THEN
    local_DesiredHeater := FALSE;
ELSIF TemperatureSensorInput < SetTemperature THEN
    local_DesiredHeater := TRUE;
ELSE
    local_DesiredHeater := FALSE;
END_IF;

HeaterOutput := local_DesiredHeater;

tmp_HeaterOnTimer(IN := HeaterOutput, PT := T#5001MS);
IF tmp_HeaterOnTimer.Q THEN
    local_OverheatActive := TRUE;
    HeaterOutput := FALSE;
END_IF;

tmp_CooldownTimer(IN := local_OverheatActive, PT := T#3S);
IF tmp_CooldownTimer.Q THEN
    local_OverheatActive := FALSE;
    IF local_SensorFault THEN
        HeaterOutput := FALSE;
    ELSIF TemperatureSensorInput < SetTemperature THEN
        HeaterOutput := TRUE;
    ELSE
        HeaterOutput := FALSE;
    END_IF;
    tmp_HeaterOnTimer(IN := HeaterOutput, PT := T#5001MS);
END_IF;

HeaterStatus := HeaterOutput;
OverheatProtection := local_OverheatActive;
END_FUNCTION_BLOCK

(* ---- public-medium-05.candidate_01.st ---- *)
(* ENGINEERING_CONTRACT
  - MotorForward/Reverse (PUB001/PUB002): manual controls selected by Mode=0; both directions inhibited on conflict.
  - MotorForward auto (PUB003/PUB004): latched start at SensorA+ButtonA or SensorB+ButtonB; reset by SensorB/SensorC; stop priority over start.
  - MotorReverse auto: forced FALSE.
  - CompletionLight (PUB004): set while Mode=1 and SensorC+ButtonC; held while SensorC=1; reset when SensorC=0.
  - Buttons are level-sensitive; no edge memory.
  - Retained latches survive mode switches; arrival resets occur even in manual.
  - BOOL arithmetic; no numeric units.
*)

(* CONTRACT_RULES [] *)

FUNCTION_BLOCK FB_ProductionLine
VAR_INPUT
    Mode : BOOL;
    ForwardButton : BOOL;
    ReverseButton : BOOL;
    SensorA : BOOL;
    SensorB : BOOL;
    SensorC : BOOL;
    ButtonA : BOOL;
    ButtonB : BOOL;
    ButtonC : BOOL;
END_VAR
VAR_OUTPUT
    MotorForward : BOOL;
    MotorReverse : BOOL;
    CompletionLight : BOOL;
END_VAR
VAR
    tmp_MoveToB : BOOL := FALSE;
    tmp_MoveToC : BOOL := FALSE;
    tmp_Completed : BOOL := FALSE;
END_VAR

// Update automatic-mode latches with stop priority.
// Movement to B starts only in automatic mode and when SensorA and ButtonA are true.
// It is cleared as soon as SensorB detects the product.
tmp_MoveToB := (tmp_MoveToB OR (Mode AND SensorA AND ButtonA)) AND NOT SensorB;

// Movement to C starts similarly from B and is cleared by SensorC.
tmp_MoveToC := (tmp_MoveToC OR (Mode AND SensorB AND ButtonB)) AND NOT SensorC;

// Completion light is set only in automatic mode when product is at C and ButtonC is pressed.
// It remains on while SensorC is true and is cleared when SensorC goes false.
tmp_Completed := (tmp_Completed OR (Mode AND SensorC AND ButtonC)) AND SensorC;

IF Mode THEN
    // Automatic mode: motor forward comes from the latched movement flags.
    MotorForward := tmp_MoveToB OR tmp_MoveToC;
    MotorReverse := FALSE;
ELSE
    // Manual mode: direct pushbutton control with interlock.
    IF ForwardButton AND NOT ReverseButton THEN
        MotorForward := TRUE;
        MotorReverse := FALSE;
    ELSIF ReverseButton AND NOT ForwardButton THEN
        MotorForward := FALSE;
        MotorReverse := TRUE;
    ELSE
        // Both or neither pressed: inhibit both directions.
        MotorForward := FALSE;
        MotorReverse := FALSE;
    END_IF;
END_IF;

// Completion light always reflects the automatic completion latch.
CompletionLight := tmp_Completed;

END_FUNCTION_BLOCK

(* ---- public-medium-05.candidate_02.st ---- *)
(* ENGINEERING_CONTRACT
  - MotorForward/Reverse (PUB001/PUB002): manual controls selected by Mode=0; both directions inhibited on conflict.
  - MotorForward auto (PUB003/PUB004): latched start at SensorA+ButtonA or SensorB+ButtonB; reset by SensorB/SensorC; stop priority over start.
  - MotorReverse auto: forced FALSE.
  - CompletionLight (PUB004): set while Mode=1 and SensorC+ButtonC; held while SensorC=1; reset when SensorC=0.
  - Automatic buttons are edge-triggered; manual direction buttons remain level.
  - Retained latches survive mode switches; arrival resets occur even in manual.
  - BOOL arithmetic; no numeric units.
*)

(* CONTRACT_RULES [] *)

FUNCTION_BLOCK FB_ProductionLine
VAR_INPUT
    Mode : BOOL;
    ForwardButton : BOOL;
    ReverseButton : BOOL;
    SensorA : BOOL;
    SensorB : BOOL;
    SensorC : BOOL;
    ButtonA : BOOL;
    ButtonB : BOOL;
    ButtonC : BOOL;
END_VAR
VAR_OUTPUT
    MotorForward : BOOL;
    MotorReverse : BOOL;
    CompletionLight : BOOL;
END_VAR
VAR
    tmp_MoveToB : BOOL := FALSE;
    tmp_MoveToC : BOOL := FALSE;
    tmp_Completed : BOOL := FALSE;
    tmp_TrigA : R_TRIG;
    tmp_TrigB : R_TRIG;
    tmp_TrigC : R_TRIG;
END_VAR

tmp_TrigA(CLK := ButtonA);
tmp_TrigB(CLK := ButtonB);
tmp_TrigC(CLK := ButtonC);

// Update automatic-mode latches with stop priority.
// Automatic commands require a rising edge on the matching button while the product sensor is true.
// Movement to B starts on a ButtonA edge with SensorA true and clears when SensorB detects the product.
tmp_MoveToB := (tmp_MoveToB OR (Mode AND SensorA AND tmp_TrigA.Q)) AND NOT SensorB;

// Movement to C starts on a ButtonB edge with SensorB true and clears when SensorC detects the product.
tmp_MoveToC := (tmp_MoveToC OR (Mode AND SensorB AND tmp_TrigB.Q)) AND NOT SensorC;

// Completion light is set on a ButtonC edge with SensorC true and remains on while SensorC is true.
// It clears as soon as the product is removed from SensorC.
tmp_Completed := (tmp_Completed OR (Mode AND SensorC AND tmp_TrigC.Q)) AND SensorC;

IF Mode THEN
    // Automatic mode: motor forward comes from the latched movement flags.
    MotorForward := tmp_MoveToB OR tmp_MoveToC;
    MotorReverse := FALSE;
ELSE
    // Manual mode: direct pushbutton control with interlock.
    IF ForwardButton AND NOT ReverseButton THEN
        MotorForward := TRUE;
        MotorReverse := FALSE;
    ELSIF ReverseButton AND NOT ForwardButton THEN
        MotorForward := FALSE;
        MotorReverse := TRUE;
    ELSE
        // Both or neither pressed: inhibit both directions.
        MotorForward := FALSE;
        MotorReverse := FALSE;
    END_IF;
END_IF;

// Completion light always reflects the automatic completion latch.
CompletionLight := tmp_Completed;

END_FUNCTION_BLOCK

(* ---- public-medium-05.candidate_03.st ---- *)
(* ENGINEERING_CONTRACT
  - MotorForward/Reverse (PUB001/PUB002): manual controls selected by Mode=0; both directions inhibited on conflict.
  - MotorForward auto (PUB003/PUB004): latched start at SensorA+ButtonA or SensorB+ButtonB; reset by SensorB/SensorC; stop priority over start.
  - MotorReverse auto: forced FALSE.
  - CompletionLight (PUB004): set while Mode=1 and SensorC+ButtonC; held while SensorC=1; reset when SensorC=0.
  - Buttons are level-sensitive; no edge memory.
  - Retained latches survive mode switches; arrival resets occur even in manual.
  - BOOL arithmetic; no numeric units.
*)

(* CONTRACT_RULES [] *)

FUNCTION_BLOCK FB_ProductionLine
VAR_INPUT
    Mode : BOOL;
    ForwardButton : BOOL;
    ReverseButton : BOOL;
    SensorA : BOOL;
    SensorB : BOOL;
    SensorC : BOOL;
    ButtonA : BOOL;
    ButtonB : BOOL;
    ButtonC : BOOL;
END_VAR
VAR_OUTPUT
    MotorForward : BOOL;
    MotorReverse : BOOL;
    CompletionLight : BOOL;
END_VAR
VAR
    tmp_MoveToB : BOOL := FALSE;
    tmp_MoveToC : BOOL := FALSE;
    tmp_Completed : BOOL := FALSE;
END_VAR

// Update automatic-mode latches with stop priority.
// Movement to B starts only in automatic mode and when SensorA and ButtonA are true.
// It is cleared as soon as SensorB detects the product.
tmp_MoveToB := (tmp_MoveToB OR (Mode AND SensorA AND ButtonA)) AND NOT SensorB;

// Movement to C starts similarly from B and is cleared by SensorC.
tmp_MoveToC := (tmp_MoveToC OR (Mode AND SensorB AND ButtonB)) AND NOT SensorC;

// Completion light is set only in automatic mode when product is at C and ButtonC is pressed.
// It remains on while SensorC is true and is cleared when SensorC goes false.
tmp_Completed := (tmp_Completed OR (Mode AND SensorC AND ButtonC)) AND SensorC;

IF Mode THEN
    // Automatic mode: motor forward comes from the latched movement flags.
    MotorForward := tmp_MoveToB OR tmp_MoveToC;
    MotorReverse := FALSE;
ELSE
    // Manual mode: clear any retained automatic sequence state.
    tmp_MoveToB := FALSE;
    tmp_MoveToC := FALSE;
    tmp_Completed := FALSE;

    // Manual mode: direct pushbutton control with interlock.
    IF ForwardButton AND NOT ReverseButton THEN
        MotorForward := TRUE;
        MotorReverse := FALSE;
    ELSIF ReverseButton AND NOT ForwardButton THEN
        MotorForward := FALSE;
        MotorReverse := TRUE;
    ELSE
        // Both or neither pressed: inhibit both directions.
        MotorForward := FALSE;
        MotorReverse := FALSE;
    END_IF;
END_IF;

// Completion light always reflects the automatic completion latch.
CompletionLight := Mode AND tmp_Completed;

END_FUNCTION_BLOCK

(* ---- public-medium-05.candidate_04.st ---- *)
(* ENGINEERING_CONTRACT
  - MotorForward/Reverse (PUB001/PUB002): manual controls selected by Mode=0; both directions inhibited on conflict.
  - MotorForward auto (PUB003/PUB004): latched start at SensorA+ButtonA or SensorB+ButtonB; reset by SensorB/SensorC; stop priority over start.
  - MotorReverse auto: forced FALSE.
  - CompletionLight (PUB004): set while Mode=1 and SensorC+ButtonC; held while SensorC=1; reset when SensorC=0.
  - Buttons are level-sensitive; no edge memory.
  - Movement latches are cleared in manual mode; completion latch survives mode switches while SensorC=1.
  - BOOL arithmetic; no numeric units.
*)

(* CONTRACT_RULES [] *)

FUNCTION_BLOCK FB_ProductionLine
VAR_INPUT
    Mode : BOOL;
    ForwardButton : BOOL;
    ReverseButton : BOOL;
    SensorA : BOOL;
    SensorB : BOOL;
    SensorC : BOOL;
    ButtonA : BOOL;
    ButtonB : BOOL;
    ButtonC : BOOL;
END_VAR
VAR_OUTPUT
    MotorForward : BOOL;
    MotorReverse : BOOL;
    CompletionLight : BOOL;
END_VAR
VAR
    tmp_MoveToB : BOOL := FALSE;
    tmp_MoveToC : BOOL := FALSE;
    tmp_Completed : BOOL := FALSE;
END_VAR

// Update automatic-mode latches with stop priority.
// Movement to B starts only in automatic mode and when SensorA and ButtonA are true.
// It is cleared as soon as SensorB detects the product.
tmp_MoveToB := (tmp_MoveToB OR (Mode AND SensorA AND ButtonA)) AND NOT SensorB;

// Movement to C starts similarly from B and is cleared by SensorC.
tmp_MoveToC := (tmp_MoveToC OR (Mode AND SensorB AND ButtonB)) AND NOT SensorC;

// Completion light is set only in automatic mode when product is at C and ButtonC is pressed.
// It remains on while SensorC is true and is cleared when SensorC goes false.
tmp_Completed := (tmp_Completed OR (Mode AND SensorC AND ButtonC)) AND SensorC;

IF Mode THEN
    // Automatic mode: motor forward comes from the latched movement flags.
    MotorForward := tmp_MoveToB OR tmp_MoveToC;
    MotorReverse := FALSE;
ELSE
    // Manual mode: movement automatic sequence state is cleared,
    // but the completion latch is retained so CompletionLight can
    // remain on until SensorC releases the product.
    tmp_MoveToB := FALSE;
    tmp_MoveToC := FALSE;

    // Manual mode: direct pushbutton control with interlock.
    IF ForwardButton AND NOT ReverseButton THEN
        MotorForward := TRUE;
        MotorReverse := FALSE;
    ELSIF ReverseButton AND NOT ForwardButton THEN
        MotorForward := FALSE;
        MotorReverse := TRUE;
    ELSE
        // Both or neither pressed: inhibit both directions.
        MotorForward := FALSE;
        MotorReverse := FALSE;
    END_IF;
END_IF;

// Completion light always reflects the automatic completion latch.
CompletionLight := tmp_Completed;

END_FUNCTION_BLOCK

(* ---- public-medium-05.patch_base_02.st ---- *)
(* ENGINEERING_CONTRACT
  - MotorForward/Reverse (PUB001/PUB002): manual controls selected by Mode=0; both directions inhibited on conflict.
  - MotorForward auto (PUB003/PUB004): latched start at SensorA+ButtonA or SensorB+ButtonB; reset by SensorB/SensorC; stop priority over start.
  - MotorReverse auto: forced FALSE.
  - CompletionLight (PUB004): set while Mode=1 and SensorC+ButtonC; held while SensorC=1; reset when SensorC=0.
  - Buttons are level-sensitive; no edge memory.
  - Retained latches survive mode switches; arrival resets occur even in manual.
  - BOOL arithmetic; no numeric units.
*)

(* CONTRACT_RULES [] *)

FUNCTION_BLOCK FB_ProductionLine
VAR_INPUT
    Mode : BOOL;
    ForwardButton : BOOL;
    ReverseButton : BOOL;
    SensorA : BOOL;
    SensorB : BOOL;
    SensorC : BOOL;
    ButtonA : BOOL;
    ButtonB : BOOL;
    ButtonC : BOOL;
END_VAR
VAR_OUTPUT
    MotorForward : BOOL;
    MotorReverse : BOOL;
    CompletionLight : BOOL;
END_VAR
VAR
    tmp_MoveToB : BOOL := FALSE;
    tmp_MoveToC : BOOL := FALSE;
    tmp_Completed : BOOL := FALSE;
END_VAR

// Update automatic-mode latches with stop priority.
// Movement to B starts only in automatic mode and when SensorA and ButtonA are true.
// It is cleared as soon as SensorB detects the product.
tmp_MoveToB := (tmp_MoveToB OR (Mode AND SensorA AND ButtonA)) AND NOT SensorB;

// Movement to C starts similarly from B and is cleared by SensorC.
tmp_MoveToC := (tmp_MoveToC OR (Mode AND SensorB AND ButtonB)) AND NOT SensorC;

// Completion light is set only in automatic mode when product is at C and ButtonC is pressed.
// It remains on while SensorC is true and is cleared when SensorC goes false.
tmp_Completed := (tmp_Completed OR (Mode AND SensorC AND ButtonC)) AND SensorC;

IF Mode THEN
    // Automatic mode: motor forward comes from the latched movement flags.
    MotorForward := tmp_MoveToB OR tmp_MoveToC;
    MotorReverse := FALSE;
ELSE
    // Manual mode: direct pushbutton control with interlock.
    IF ForwardButton AND NOT ReverseButton THEN
        MotorForward := TRUE;
        MotorReverse := FALSE;
    ELSIF ReverseButton AND NOT ForwardButton THEN
        MotorForward := FALSE;
        MotorReverse := TRUE;
    ELSE
        // Both or neither pressed: inhibit both directions.
        MotorForward := FALSE;
        MotorReverse := FALSE;
    END_IF;
END_IF;

// Completion light always reflects the automatic completion latch.
CompletionLight := tmp_Completed;

END_FUNCTION_BLOCK

(* ---- public-medium-05.patch_base_03.st ---- *)
(* ENGINEERING_CONTRACT
  - MotorForward/Reverse (PUB001/PUB002): manual controls selected by Mode=0; both directions inhibited on conflict.
  - MotorForward auto (PUB003/PUB004): latched start at SensorA+ButtonA or SensorB+ButtonB; reset by SensorB/SensorC; stop priority over start.
  - MotorReverse auto: forced FALSE.
  - CompletionLight (PUB004): set while Mode=1 and SensorC+ButtonC; held while SensorC=1; reset when SensorC=0.
  - Buttons are level-sensitive; no edge memory.
  - Retained latches survive mode switches; arrival resets occur even in manual.
  - BOOL arithmetic; no numeric units.
*)

(* CONTRACT_RULES [] *)

FUNCTION_BLOCK FB_ProductionLine
VAR_INPUT
    Mode : BOOL;
    ForwardButton : BOOL;
    ReverseButton : BOOL;
    SensorA : BOOL;
    SensorB : BOOL;
    SensorC : BOOL;
    ButtonA : BOOL;
    ButtonB : BOOL;
    ButtonC : BOOL;
END_VAR
VAR_OUTPUT
    MotorForward : BOOL;
    MotorReverse : BOOL;
    CompletionLight : BOOL;
END_VAR
VAR
    tmp_MoveToB : BOOL := FALSE;
    tmp_MoveToC : BOOL := FALSE;
    tmp_Completed : BOOL := FALSE;
END_VAR

// Update automatic-mode latches with stop priority.
// Movement to B starts only in automatic mode and when SensorA and ButtonA are true.
// It is cleared as soon as SensorB detects the product.
tmp_MoveToB := (tmp_MoveToB OR (Mode AND SensorA AND ButtonA)) AND NOT SensorB;

// Movement to C starts similarly from B and is cleared by SensorC.
tmp_MoveToC := (tmp_MoveToC OR (Mode AND SensorB AND ButtonB)) AND NOT SensorC;

// Completion light is set only in automatic mode when product is at C and ButtonC is pressed.
// It remains on while SensorC is true and is cleared when SensorC goes false.
tmp_Completed := (tmp_Completed OR (Mode AND SensorC AND ButtonC)) AND SensorC;

IF Mode THEN
    // Automatic mode: motor forward comes from the latched movement flags.
    MotorForward := tmp_MoveToB OR tmp_MoveToC;
    MotorReverse := FALSE;
ELSE
    // Manual mode: direct pushbutton control with interlock.
    IF ForwardButton AND NOT ReverseButton THEN
        MotorForward := TRUE;
        MotorReverse := FALSE;
    ELSIF ReverseButton AND NOT ForwardButton THEN
        MotorForward := FALSE;
        MotorReverse := TRUE;
    ELSE
        // Both or neither pressed: inhibit both directions.
        MotorForward := FALSE;
        MotorReverse := FALSE;
    END_IF;
END_IF;

// Completion light always reflects the automatic completion latch.
CompletionLight := tmp_Completed;

END_FUNCTION_BLOCK

(* ---- public-medium-05.patch_base_04.st ---- *)
(* ENGINEERING_CONTRACT
  - MotorForward/Reverse (PUB001/PUB002): manual controls selected by Mode=0; both directions inhibited on conflict.
  - MotorForward auto (PUB003/PUB004): latched start at SensorA+ButtonA or SensorB+ButtonB; reset by SensorB/SensorC; stop priority over start.
  - MotorReverse auto: forced FALSE.
  - CompletionLight (PUB004): set while Mode=1 and SensorC+ButtonC; held while SensorC=1; reset when SensorC=0.
  - Buttons are level-sensitive; no edge memory.
  - Retained latches survive mode switches; arrival resets occur even in manual.
  - BOOL arithmetic; no numeric units.
*)

(* CONTRACT_RULES [] *)

FUNCTION_BLOCK FB_ProductionLine
VAR_INPUT
    Mode : BOOL;
    ForwardButton : BOOL;
    ReverseButton : BOOL;
    SensorA : BOOL;
    SensorB : BOOL;
    SensorC : BOOL;
    ButtonA : BOOL;
    ButtonB : BOOL;
    ButtonC : BOOL;
END_VAR
VAR_OUTPUT
    MotorForward : BOOL;
    MotorReverse : BOOL;
    CompletionLight : BOOL;
END_VAR
VAR
    tmp_MoveToB : BOOL := FALSE;
    tmp_MoveToC : BOOL := FALSE;
    tmp_Completed : BOOL := FALSE;
END_VAR

// Update automatic-mode latches with stop priority.
// Movement to B starts only in automatic mode and when SensorA and ButtonA are true.
// It is cleared as soon as SensorB detects the product.
tmp_MoveToB := (tmp_MoveToB OR (Mode AND SensorA AND ButtonA)) AND NOT SensorB;

// Movement to C starts similarly from B and is cleared by SensorC.
tmp_MoveToC := (tmp_MoveToC OR (Mode AND SensorB AND ButtonB)) AND NOT SensorC;

// Completion light is set only in automatic mode when product is at C and ButtonC is pressed.
// It remains on while SensorC is true and is cleared when SensorC goes false.
tmp_Completed := (tmp_Completed OR (Mode AND SensorC AND ButtonC)) AND SensorC;

IF Mode THEN
    // Automatic mode: motor forward comes from the latched movement flags.
    MotorForward := tmp_MoveToB OR tmp_MoveToC;
    MotorReverse := FALSE;
ELSE
    // Manual mode: clear any retained automatic sequence state.
    tmp_MoveToB := FALSE;
    tmp_MoveToC := FALSE;
    tmp_Completed := FALSE;

    // Manual mode: direct pushbutton control with interlock.
    IF ForwardButton AND NOT ReverseButton THEN
        MotorForward := TRUE;
        MotorReverse := FALSE;
    ELSIF ReverseButton AND NOT ForwardButton THEN
        MotorForward := FALSE;
        MotorReverse := TRUE;
    ELSE
        // Both or neither pressed: inhibit both directions.
        MotorForward := FALSE;
        MotorReverse := FALSE;
    END_IF;
END_IF;

// Completion light always reflects the automatic completion latch.
CompletionLight := Mode AND tmp_Completed;

END_FUNCTION_BLOCK

(* ---- public-medium-05.raw_candidate_01.st ---- *)
(* ENGINEERING_CONTRACT
  - MotorForward/Reverse (PUB001/PUB002): manual controls selected by Mode=0; both directions inhibited on conflict.
  - MotorForward auto (PUB003/PUB004): latched start at SensorA+ButtonA or SensorB+ButtonB; reset by SensorB/SensorC; stop priority over start.
  - MotorReverse auto: forced FALSE.
  - CompletionLight (PUB004): set while Mode=1 and SensorC+ButtonC; held while SensorC=1; reset when SensorC=0.
  - Buttons are level-sensitive; no edge memory.
  - Retained latches survive mode switches; arrival resets occur even in manual.
  - BOOL arithmetic; no numeric units.
*)

(* CONTRACT_RULES [] *)

FUNCTION_BLOCK FB_ProductionLine
VAR_INPUT
    Mode : BOOL;
    ForwardButton : BOOL;
    ReverseButton : BOOL;
    SensorA : BOOL;
    SensorB : BOOL;
    SensorC : BOOL;
    ButtonA : BOOL;
    ButtonB : BOOL;
    ButtonC : BOOL;
END_VAR
VAR_OUTPUT
    MotorForward : BOOL;
    MotorReverse : BOOL;
    CompletionLight : BOOL;
END_VAR
VAR
    tmp_MoveToB : BOOL := FALSE;
    tmp_MoveToC : BOOL := FALSE;
    tmp_Completed : BOOL := FALSE;
END_VAR

// Update automatic-mode latches with stop priority.
// Movement to B starts only in automatic mode and when SensorA and ButtonA are true.
// It is cleared as soon as SensorB detects the product.
tmp_MoveToB := (tmp_MoveToB OR (Mode AND SensorA AND ButtonA)) AND NOT SensorB;

// Movement to C starts similarly from B and is cleared by SensorC.
tmp_MoveToC := (tmp_MoveToC OR (Mode AND SensorB AND ButtonB)) AND NOT SensorC;

// Completion light is set only in automatic mode when product is at C and ButtonC is pressed.
// It remains on while SensorC is true and is cleared when SensorC goes false.
tmp_Completed := (tmp_Completed OR (Mode AND SensorC AND ButtonC)) AND SensorC;

IF Mode THEN
    // Automatic mode: motor forward comes from the latched movement flags.
    MotorForward := tmp_MoveToB OR tmp_MoveToC;
    MotorReverse := FALSE;
ELSE
    // Manual mode: direct pushbutton control with interlock.
    IF ForwardButton AND NOT ReverseButton THEN
        MotorForward := TRUE;
        MotorReverse := FALSE;
    ELSIF ReverseButton AND NOT ForwardButton THEN
        MotorForward := FALSE;
        MotorReverse := TRUE;
    ELSE
        // Both or neither pressed: inhibit both directions.
        MotorForward := FALSE;
        MotorReverse := FALSE;
    END_IF;
END_IF;

// Completion light always reflects the automatic completion latch.
CompletionLight := tmp_Completed;

END_FUNCTION_BLOCK

(* ---- public-medium-05.raw_candidate_02.st ---- *)
(* ENGINEERING_CONTRACT
  - MotorForward/Reverse (PUB001/PUB002): manual controls selected by Mode=0; both directions inhibited on conflict.
  - MotorForward auto (PUB003/PUB004): latched start at SensorA+ButtonA or SensorB+ButtonB; reset by SensorB/SensorC; stop priority over start.
  - MotorReverse auto: forced FALSE.
  - CompletionLight (PUB004): set while Mode=1 and SensorC+ButtonC; held while SensorC=1; reset when SensorC=0.
  - Automatic buttons are edge-triggered; manual direction buttons remain level.
  - Retained latches survive mode switches; arrival resets occur even in manual.
  - BOOL arithmetic; no numeric units.
*)

(* CONTRACT_RULES [] *)

FUNCTION_BLOCK FB_ProductionLine
VAR_INPUT
    Mode : BOOL;
    ForwardButton : BOOL;
    ReverseButton : BOOL;
    SensorA : BOOL;
    SensorB : BOOL;
    SensorC : BOOL;
    ButtonA : BOOL;
    ButtonB : BOOL;
    ButtonC : BOOL;
END_VAR
VAR_OUTPUT
    MotorForward : BOOL;
    MotorReverse : BOOL;
    CompletionLight : BOOL;
END_VAR
VAR
    tmp_MoveToB : BOOL := FALSE;
    tmp_MoveToC : BOOL := FALSE;
    tmp_Completed : BOOL := FALSE;
    tmp_TrigA : R_TRIG;
    tmp_TrigB : R_TRIG;
    tmp_TrigC : R_TRIG;
END_VAR

tmp_TrigA(CLK := ButtonA);
tmp_TrigB(CLK := ButtonB);
tmp_TrigC(CLK := ButtonC);

// Update automatic-mode latches with stop priority.
// Automatic commands require a rising edge on the matching button while the product sensor is true.
// Movement to B starts on a ButtonA edge with SensorA true and clears when SensorB detects the product.
tmp_MoveToB := (tmp_MoveToB OR (Mode AND SensorA AND tmp_TrigA.Q)) AND NOT SensorB;

// Movement to C starts on a ButtonB edge with SensorB true and clears when SensorC detects the product.
tmp_MoveToC := (tmp_MoveToC OR (Mode AND SensorB AND tmp_TrigB.Q)) AND NOT SensorC;

// Completion light is set on a ButtonC edge with SensorC true and remains on while SensorC is true.
// It clears as soon as the product is removed from SensorC.
tmp_Completed := (tmp_Completed OR (Mode AND SensorC AND tmp_TrigC.Q)) AND SensorC;

IF Mode THEN
    // Automatic mode: motor forward comes from the latched movement flags.
    MotorForward := tmp_MoveToB OR tmp_MoveToC;
    MotorReverse := FALSE;
ELSE
    // Manual mode: direct pushbutton control with interlock.
    IF ForwardButton AND NOT ReverseButton THEN
        MotorForward := TRUE;
        MotorReverse := FALSE;
    ELSIF ReverseButton AND NOT ForwardButton THEN
        MotorForward := FALSE;
        MotorReverse := TRUE;
    ELSE
        // Both or neither pressed: inhibit both directions.
        MotorForward := FALSE;
        MotorReverse := FALSE;
    END_IF;
END_IF;

// Completion light always reflects the automatic completion latch.
CompletionLight := tmp_Completed;

END_FUNCTION_BLOCK

(* ---- public-medium-05.raw_candidate_03.st ---- *)
(* ENGINEERING_CONTRACT
  - MotorForward/Reverse (PUB001/PUB002): manual controls selected by Mode=0; both directions inhibited on conflict.
  - MotorForward auto (PUB003/PUB004): latched start at SensorA+ButtonA or SensorB+ButtonB; reset by SensorB/SensorC; stop priority over start.
  - MotorReverse auto: forced FALSE.
  - CompletionLight (PUB004): set while Mode=1 and SensorC+ButtonC; held while SensorC=1; reset when SensorC=0.
  - Buttons are level-sensitive; no edge memory.
  - Retained latches survive mode switches; arrival resets occur even in manual.
  - BOOL arithmetic; no numeric units.
*)

(* CONTRACT_RULES [] *)

FUNCTION_BLOCK FB_ProductionLine
VAR_INPUT
    Mode : BOOL;
    ForwardButton : BOOL;
    ReverseButton : BOOL;
    SensorA : BOOL;
    SensorB : BOOL;
    SensorC : BOOL;
    ButtonA : BOOL;
    ButtonB : BOOL;
    ButtonC : BOOL;
END_VAR
VAR_OUTPUT
    MotorForward : BOOL;
    MotorReverse : BOOL;
    CompletionLight : BOOL;
END_VAR
VAR
    tmp_MoveToB : BOOL := FALSE;
    tmp_MoveToC : BOOL := FALSE;
    tmp_Completed : BOOL := FALSE;
END_VAR

// Update automatic-mode latches with stop priority.
// Movement to B starts only in automatic mode and when SensorA and ButtonA are true.
// It is cleared as soon as SensorB detects the product.
tmp_MoveToB := (tmp_MoveToB OR (Mode AND SensorA AND ButtonA)) AND NOT SensorB;

// Movement to C starts similarly from B and is cleared by SensorC.
tmp_MoveToC := (tmp_MoveToC OR (Mode AND SensorB AND ButtonB)) AND NOT SensorC;

// Completion light is set only in automatic mode when product is at C and ButtonC is pressed.
// It remains on while SensorC is true and is cleared when SensorC goes false.
tmp_Completed := (tmp_Completed OR (Mode AND SensorC AND ButtonC)) AND SensorC;

IF Mode THEN
    // Automatic mode: motor forward comes from the latched movement flags.
    MotorForward := tmp_MoveToB OR tmp_MoveToC;
    MotorReverse := FALSE;
ELSE
    // Manual mode: clear any retained automatic sequence state.
    tmp_MoveToB := FALSE;
    tmp_MoveToC := FALSE;
    tmp_Completed := FALSE;

    // Manual mode: direct pushbutton control with interlock.
    IF ForwardButton AND NOT ReverseButton THEN
        MotorForward := TRUE;
        MotorReverse := FALSE;
    ELSIF ReverseButton AND NOT ForwardButton THEN
        MotorForward := FALSE;
        MotorReverse := TRUE;
    ELSE
        // Both or neither pressed: inhibit both directions.
        MotorForward := FALSE;
        MotorReverse := FALSE;
    END_IF;
END_IF;

// Completion light always reflects the automatic completion latch.
CompletionLight := Mode AND tmp_Completed;

END_FUNCTION_BLOCK

(* ---- public-medium-05.raw_candidate_04.st ---- *)
(* ENGINEERING_CONTRACT
  - MotorForward/Reverse (PUB001/PUB002): manual controls selected by Mode=0; both directions inhibited on conflict.
  - MotorForward auto (PUB003/PUB004): latched start at SensorA+ButtonA or SensorB+ButtonB; reset by SensorB/SensorC; stop priority over start.
  - MotorReverse auto: forced FALSE.
  - CompletionLight (PUB004): set while Mode=1 and SensorC+ButtonC; held while SensorC=1; reset when SensorC=0.
  - Buttons are level-sensitive; no edge memory.
  - Movement latches are cleared in manual mode; completion latch survives mode switches while SensorC=1.
  - BOOL arithmetic; no numeric units.
*)

(* CONTRACT_RULES [] *)

FUNCTION_BLOCK FB_ProductionLine
VAR_INPUT
    Mode : BOOL;
    ForwardButton : BOOL;
    ReverseButton : BOOL;
    SensorA : BOOL;
    SensorB : BOOL;
    SensorC : BOOL;
    ButtonA : BOOL;
    ButtonB : BOOL;
    ButtonC : BOOL;
END_VAR
VAR_OUTPUT
    MotorForward : BOOL;
    MotorReverse : BOOL;
    CompletionLight : BOOL;
END_VAR
VAR
    tmp_MoveToB : BOOL := FALSE;
    tmp_MoveToC : BOOL := FALSE;
    tmp_Completed : BOOL := FALSE;
END_VAR

// Update automatic-mode latches with stop priority.
// Movement to B starts only in automatic mode and when SensorA and ButtonA are true.
// It is cleared as soon as SensorB detects the product.
tmp_MoveToB := (tmp_MoveToB OR (Mode AND SensorA AND ButtonA)) AND NOT SensorB;

// Movement to C starts similarly from B and is cleared by SensorC.
tmp_MoveToC := (tmp_MoveToC OR (Mode AND SensorB AND ButtonB)) AND NOT SensorC;

// Completion light is set only in automatic mode when product is at C and ButtonC is pressed.
// It remains on while SensorC is true and is cleared when SensorC goes false.
tmp_Completed := (tmp_Completed OR (Mode AND SensorC AND ButtonC)) AND SensorC;

IF Mode THEN
    // Automatic mode: motor forward comes from the latched movement flags.
    MotorForward := tmp_MoveToB OR tmp_MoveToC;
    MotorReverse := FALSE;
ELSE
    // Manual mode: movement automatic sequence state is cleared,
    // but the completion latch is retained so CompletionLight can
    // remain on until SensorC releases the product.
    tmp_MoveToB := FALSE;
    tmp_MoveToC := FALSE;

    // Manual mode: direct pushbutton control with interlock.
    IF ForwardButton AND NOT ReverseButton THEN
        MotorForward := TRUE;
        MotorReverse := FALSE;
    ELSIF ReverseButton AND NOT ForwardButton THEN
        MotorForward := FALSE;
        MotorReverse := TRUE;
    ELSE
        // Both or neither pressed: inhibit both directions.
        MotorForward := FALSE;
        MotorReverse := FALSE;
    END_IF;
END_IF;

// Completion light always reflects the automatic completion latch.
CompletionLight := tmp_Completed;

END_FUNCTION_BLOCK

(* ---- public-medium-07.candidate_01.st ---- *)
(* CONTRACT_RULES [] *)
(* ENGINEERING_CONTRACT
Group | Activation | Retention | Reset | Same-scan priority | Units/boundaries
SUPPLY_FAN_RUN | enable=OCCUPANCY_DETECTED AND HVAC_MODE_SELECTOR<>3 for T#30S continuously | TON holds Q true while enable true and elapsed>=PT | IN false clears ET and Q on same call | timer called before Q copied | BOOL, seconds (PUB002,PUB007)
TEMP_SETPOINT_ADJUST | valid mode combinational from current inputs | none; recomputed each scan | next input scan overwrites | clamp after raw calculation | INT degC, [-4,4] (PUB003-PUB006)
*)
FUNCTION_BLOCK OfficeHVACControl
VAR_INPUT
    OCCUPANCY_DETECTED : BOOL;
    ENERGY_SAVING_MODE : BOOL;
    HVAC_MODE_SELECTOR : INT;
END_VAR
VAR_OUTPUT
    SUPPLY_FAN_RUN : BOOL;
    TEMP_SETPOINT_ADJUST : INT;
END_VAR
VAR
    local_fan_timer : TON;
    local_fan_enable : BOOL;
    local_raw_adjust : INT;
END_VAR

local_fan_enable := OCCUPANCY_DETECTED AND (HVAC_MODE_SELECTOR <> 3);
local_fan_timer(IN := local_fan_enable, PT := T#30S);
SUPPLY_FAN_RUN := local_fan_timer.Q;

CASE HVAC_MODE_SELECTOR OF
    0:
        IF OCCUPANCY_DETECTED THEN
            local_raw_adjust := 0;
        ELSIF ENERGY_SAVING_MODE THEN
            local_raw_adjust := 3;
        ELSE
            local_raw_adjust := 2;
        END_IF;
    1:
        IF OCCUPANCY_DETECTED THEN
            local_raw_adjust := 0;
        ELSE
            local_raw_adjust := 1;
        END_IF;
    2:
        IF OCCUPANCY_DETECTED THEN
            local_raw_adjust := 0;
        ELSE
            local_raw_adjust := 4;
        END_IF;
    3:
        local_raw_adjust := 4;
    ELSE
        local_raw_adjust := 0;
END_CASE;

IF local_raw_adjust < -4 THEN
    TEMP_SETPOINT_ADJUST := -4;
ELSIF local_raw_adjust > 4 THEN
    TEMP_SETPOINT_ADJUST := 4;
ELSE
    TEMP_SETPOINT_ADJUST := local_raw_adjust;
END_IF;

END_FUNCTION_BLOCK

(* ---- public-medium-07.raw_candidate_01.st ---- *)
(* CONTRACT_RULES [] *)
(* ENGINEERING_CONTRACT
Group | Activation | Retention | Reset | Same-scan priority | Units/boundaries
SUPPLY_FAN_RUN | enable=OCCUPANCY_DETECTED AND HVAC_MODE_SELECTOR<>3 for T#30S continuously | TON holds Q true while enable true and elapsed>=PT | IN false clears ET and Q on same call | timer called before Q copied | BOOL, seconds (PUB002,PUB007)
TEMP_SETPOINT_ADJUST | valid mode combinational from current inputs | none; recomputed each scan | next input scan overwrites | clamp after raw calculation | INT degC, [-4,4] (PUB003-PUB006)
*)
FUNCTION_BLOCK OfficeHVACControl
VAR_INPUT
    OCCUPANCY_DETECTED : BOOL;
    ENERGY_SAVING_MODE : BOOL;
    HVAC_MODE_SELECTOR : INT;
END_VAR
VAR_OUTPUT
    SUPPLY_FAN_RUN : BOOL;
    TEMP_SETPOINT_ADJUST : INT;
END_VAR
VAR
    local_fan_timer : TON;
    local_fan_enable : BOOL;
    local_raw_adjust : INT;
END_VAR

local_fan_enable := OCCUPANCY_DETECTED AND (HVAC_MODE_SELECTOR <> 3);
local_fan_timer(IN := local_fan_enable, PT := T#30S);
SUPPLY_FAN_RUN := local_fan_timer.Q;

CASE HVAC_MODE_SELECTOR OF
    0:
        IF OCCUPANCY_DETECTED THEN
            local_raw_adjust := 0;
        ELSIF ENERGY_SAVING_MODE THEN
            local_raw_adjust := 3;
        ELSE
            local_raw_adjust := 2;
        END_IF;
    1:
        IF OCCUPANCY_DETECTED THEN
            local_raw_adjust := 0;
        ELSE
            local_raw_adjust := 1;
        END_IF;
    2:
        IF OCCUPANCY_DETECTED THEN
            local_raw_adjust := 0;
        ELSE
            local_raw_adjust := 4;
        END_IF;
    3:
        local_raw_adjust := 4;
    ELSE
        local_raw_adjust := 0;
END_CASE;

IF local_raw_adjust < -4 THEN
    TEMP_SETPOINT_ADJUST := -4;
ELSIF local_raw_adjust > 4 THEN
    TEMP_SETPOINT_ADJUST := 4;
ELSE
    TEMP_SETPOINT_ADJUST := local_raw_adjust;
END_IF;

END_FUNCTION_BLOCK

(* ---- public-medium-08.candidate_01.st ---- *)
FUNCTION_BLOCK IPv4Parser
(* ENGINEERING_CONTRACT
   Output ipValue: combinational UDINT, written every invocation from current ipText.
   Activation: all four segments valid (PUB001-PUB004). Retention: none; invalid sets 0 same scan.
   Reset: malformed/nondigit/incorrect count/out-of-range sets 0 (PUB001/PUB002/PUB003).
   Same-scan priority: final parse result only; no latches.
   Units/boundaries: network byte order UDINT, first octet bits 31..24, fourth octet bits 7..0; each octet 0..255.
*)
(* CONTRACT_RULES [] *)
VAR_INPUT
    ipText : STRING(254);
END_VAR
VAR_OUTPUT
    ipValue : UDINT;
END_VAR
VAR
    tmp_len : INT;
    tmp_i : INT;
    tmp_c : BYTE;
    tmp_digit : INT;
    tmp_val : UDINT;
    tmp_digits_in_seg : INT;
    tmp_seg_count : INT;
    tmp_ok : BOOL;
    tmp_result : UDINT;
END_VAR

tmp_len := LEN(ipText);

IF (tmp_len < 7) OR (tmp_len > 15) THEN
    ipValue := UDINT#0;
    RETURN;
END_IF;

tmp_i := 0;
tmp_seg_count := 0;
tmp_digits_in_seg := 0;
tmp_val := UDINT#0;
tmp_result := UDINT#0;
tmp_ok := TRUE;

WHILE (tmp_i < tmp_len) AND tmp_ok DO
    tmp_c := ipText[tmp_i];

    IF (tmp_c >= BYTE#48) AND (tmp_c <= BYTE#57) THEN
        tmp_digit := BYTE_TO_INT(tmp_c) - 48;

        IF tmp_val > UDINT#25 THEN
            tmp_ok := FALSE;
        ELSE
            tmp_val := (tmp_val * UDINT#10) + INT_TO_UDINT(tmp_digit);
            tmp_digits_in_seg := tmp_digits_in_seg + 1;
        END_IF;

    ELSIF tmp_c = BYTE#46 THEN
        IF (tmp_digits_in_seg = 0) OR (tmp_val > UDINT#255) OR (tmp_seg_count >= 3) THEN
            tmp_ok := FALSE;
        ELSE
            tmp_result := SHL(tmp_result, 8);
            tmp_result := tmp_result OR tmp_val;

            tmp_seg_count := tmp_seg_count + 1;
            tmp_val := UDINT#0;
            tmp_digits_in_seg := 0;
        END_IF;

    ELSE
        tmp_ok := FALSE;
    END_IF;

    tmp_i := tmp_i + 1;
END_WHILE;

IF tmp_ok THEN
    IF (tmp_digits_in_seg = 0) OR (tmp_val > UDINT#255) OR (tmp_seg_count <> 3) THEN
        tmp_ok := FALSE;
    END_IF;
END_IF;

IF tmp_ok THEN
    tmp_result := SHL(tmp_result, 8);
    tmp_result := tmp_result OR tmp_val;
    ipValue := tmp_result;
ELSE
    ipValue := UDINT#0;
END_IF;

END_FUNCTION_BLOCK

(* ---- public-medium-08.raw_candidate_01.st ---- *)
FUNCTION_BLOCK IPv4Parser
(* ENGINEERING_CONTRACT
   Output ipValue: combinational UDINT, written every invocation from current ipText.
   Activation: all four segments valid (PUB001-PUB004). Retention: none; invalid sets 0 same scan.
   Reset: malformed/nondigit/incorrect count/out-of-range sets 0 (PUB001/PUB002/PUB003).
   Same-scan priority: final parse result only; no latches.
   Units/boundaries: network byte order UDINT, first octet bits 31..24, fourth octet bits 7..0; each octet 0..255.
*)
(* CONTRACT_RULES [] *)
VAR_INPUT
    ipText : STRING(254);
END_VAR
VAR_OUTPUT
    ipValue : UDINT;
END_VAR
VAR
    tmp_len : INT;
    tmp_i : INT;
    tmp_c : BYTE;
    tmp_digit : INT;
    tmp_val : UDINT;
    tmp_digits_in_seg : INT;
    tmp_seg_count : INT;
    tmp_ok : BOOL;
    tmp_result : UDINT;
END_VAR

tmp_len := LEN(ipText);

IF (tmp_len < 7) OR (tmp_len > 15) THEN
    ipValue := UDINT#0;
    RETURN;
END_IF

tmp_i := 0;
tmp_seg_count := 0;
tmp_digits_in_seg := 0;
tmp_val := UDINT#0;
tmp_result := UDINT#0;
tmp_ok := TRUE;

WHILE (tmp_i < tmp_len) AND tmp_ok DO
    tmp_c := ipText[tmp_i];

    IF (tmp_c >= BYTE#48) AND (tmp_c <= BYTE#57) THEN
        tmp_digit := BYTE_TO_INT(tmp_c) - 48;

        IF tmp_val > UDINT#25 THEN
            tmp_ok := FALSE;
        ELSE
            tmp_val := (tmp_val * UDINT#10) + INT_TO_UDINT(tmp_digit);
            tmp_digits_in_seg := tmp_digits_in_seg + 1;
        END_IF;

    ELSIF tmp_c = BYTE#46 THEN
        IF (tmp_digits_in_seg = 0) OR (tmp_val > UDINT#255) OR (tmp_seg_count >= 3) THEN
            tmp_ok := FALSE;
        ELSE
            tmp_result := SHL(tmp_result, 8);
            tmp_result := tmp_result OR tmp_val;

            tmp_seg_count := tmp_seg_count + 1;
            tmp_val := UDINT#0;
            tmp_digits_in_seg := 0;
        END_IF;

    ELSE
        tmp_ok := FALSE;
    END_IF;

    tmp_i := tmp_i + 1;
END_WHILE;

IF tmp_ok THEN
    IF (tmp_digits_in_seg = 0) OR (tmp_val > UDINT#255) OR (tmp_seg_count <> 3) THEN
        tmp_ok := FALSE;
    END_IF;
END_IF;

IF tmp_ok THEN
    tmp_result := SHL(tmp_result, 8);
    tmp_result := tmp_result OR tmp_val;
    ipValue := tmp_result;
ELSE
    ipValue := UDINT#0;
END_IF;

END_FUNCTION_BLOCK
